{attribute 'Tc2GvlVarNames'}
VAR_GLOBAL
	stgGr02HMI			:ST_Gr02HMIRef;
END_VAR

(* stored: Version 1.1.0.1, ProductVersion 3.1.4024.15
   GVL GVL_Gr02HMI: Id {87aaff53-21ca-4043-8b6a-f4d9276c0c6f} *)
